PROGRAM MAIN
VAR
	
	PlcFirstCycle : BOOL := TRUE;

	// SWITCHES
	SwitchR1Up : fbSwitch;
	SwitchR1UpConfig : stSwitchConfig;
	SwitchR1Down : fbSwitch;
	SwitchR1DownConfig : stSwitchConfig;
	
	// SHUTTERS
	Shutter1 : fbShutter;
	Shutter1Cmd : stShutterCommand;
	Shutter1Config : stShutterConfig;
	
END_VAR


IF PlcFirstCycle THEN
	SwitchR1UpConfig.ShortClickMaxTime := T#500MS;
	SwitchR1UpConfig.ShortClickDelayTime := T#500MS;
	SwitchR1UpConfig.LongClickMaxTime := T#1500MS;
	
	SwitchR1DownConfig.ShortClickMaxTime := T#500MS;
	SwitchR1DownConfig.ShortClickDelayTime := T#500MS;
	SwitchR1DownConfig.LongClickMaxTime := T#1500MS;
	
	Shutter1Config.TravelTime := T#15S;
	Shutter1Config.AngleFullTurnTime := T#3S;
	
	PlcFirstCycle := FALSE;
END_IF


SwitchR1Up(I_Switch := gvlSwitches.gvSwitchR1Up, Config := SwitchR1UpConfig);
SwitchR1Down(I_Switch := gvlSwitches.gvSwitchR1Down, Config := SwitchR1DownConfig);

Shutter1Cmd.CommandType := eShutterCommandType.NONE;

// STOP condition - If shutter is moving, any switch R1 or R2 click will stop shutter
IF Shutter1.State.CurrentState <> eShutterStateType.IDLE AND 
	( SwitchR1Up.State.CurrentState <> eSwitchStateType.IDLE
	OR SwitchR1Down.State.CurrentState <> eSwitchStateType.IDLE) THEN
	Shutter1Cmd.CommandType := eShutterCommandType.STOP;

// OPEN condition
ELSIF SwitchR1Up.State.CurrentState = eSwitchStateType.MULTI_CLICK AND SwitchR1Up.State.PressCount = 2 THEN
	Shutter1Cmd.CommandType := eShutterCommandType.OPEN;

// Close condition
ELSIF SwitchR1Down.State.CurrentState = eSwitchStateType.MULTI_CLICK AND SwitchR1Down.State.PressCount = 2 THEN
	Shutter1Cmd.CommandType := eShutterCommandType.Close;

// STEP_OPEN condition
ELSIF SwitchR1Up.State.CurrentState = eSwitchStateType.SHORT_CLICK THEN
	Shutter1Cmd.CommandType := eShutterCommandType.STEP_OPEN;
	
// STEP_CLOSE condition
ELSIF SwitchR1Down.State.CurrentState = eSwitchStateType.SHORT_CLICK THEN
	Shutter1Cmd.CommandType := eShutterCommandType.STEP_CLOSE;
	
// MOVE_TO_POSITION condition
ELSIF SwitchR1Up.State.CurrentState = eSwitchStateType.LONG_CLICK
	OR SwitchR1Down.State.CurrentState = eSwitchStateType.LONG_CLICK THEN
	Shutter1Cmd.Position := 50;
	Shutter1Cmd.Angle := 50;
	Shutter1Cmd.CommandType := eShutterCommandType.MOVE_TO_POSITION;
END_IF

Shutter1(Command := Shutter1Cmd, Config := Shutter1Config);

gvlShutters.gvShutter1Up := Shutter1.Q_MoveUp;
gvlShutters.gvShutter1Down := Shutter1.Q_MoveDown;

END_PROGRAM

(* stored: Version 1.1.0.1
   POU MAIN: Id {b477ade9-5e41-44da-827a-03687596879d}, SpecialFunc None *)
